(* IEC 61131-3 sources: Lasal-MCP/examples/SampleSource/LASALScreenAdvancedSolution/LASALScreenAdvancedSolution/LASALScreenAdvacnedSolution/Stations/Terminal/HMI/Class/DragDropArea, 1 file *)

(* ---- DragDropArea.st ---- *)
(*!
<Class
	Name               = "DragDropArea"
	Revision           = "0.0"
	RealtimeTask       = "false"
	CyclicTask         = "false"
	BackgroundTask     = "false"
	Sigmatek           = "false"
	OSInterface        = "false"
	HighPriority       = "false"
	Automatic          = "false"
	UpdateMode         = "Prescan"
	SharedCommandTable = "true"
	Objectsize         = "(420,240)">
	<Channels>
		<Server Name="UpdateIcon" Visualized="false" Initialize="false" WriteProtected="false" Retentive="false"/>
		<Client Name="_Grafix" Required="false" Internal="false"/>
	</Channels>
	<Network Name="DragDropArea">
		<!-- List of Components in this network -->
		<Components>
			<Object
				Name       = "_base"
				Class      = "_MyIO"
				Position   = "(218,120)"
				Visualized = "true"
				Remotely   = "true">
				<Channels>
					<Server Name="Refresh"/>
					<Server Name="Server0"/>
					<Client Name="Graphic"/>
					<Client Name="Lse"/>
				</Channels>
			</Object>
		</Components>
		<Comments>
		</Comments>
		<!-- List of Connections in this network -->
		<Connections>
			<Connection Source="this.Server0" Destination="_base.Server0" Vertices="(706,210),(534,210),"/>
			<Connection Source="this.Refresh" Destination="_base.Refresh" Vertices="(706,270),(534,270),"/>
			<Connection Source="_base.Lse" Destination="this.Lse" Vertices="(218,210),(38,210),"/>
		</Connections>
		<!-- Headerfiles -->
		<Options>
		</Options>
	</Network>
</Class>
*)
#pragma using _MyIO

DragDropArea : CLASS
: _MyIO
  //Servers:
	UpdateIcon 	: SvrCh_DINT;
  //Clients:
	_Grafix 	: CltChCmd__Grafix;
  //Variables:
		DrawClearScreen 	: BOOL;
		Started 	: BOOL;
		OnlyOnce 	: BOOL;
		SelectedLineNo 	: DINT;
		TouchCoord 	: _DOT;
		myPio 	: _IO;
		pBMP 	: ^_BMP;
  //Functions:
				//! <Function Comment="this method is called everytime when the input is active and a event occured" Name="GetEvent"/>
	FUNCTION __CDECL VIRTUAL GLOBAL GetEvent
		VAR_INPUT
			ped 	: ^_EDITOR;			//! <Variable Comment="pointer to _EDITOR information" Name="GetEvent.ped"/>
			pe 	: ^_EVENT;			//! <Variable Comment="pointer to _EVENT information" Name="GetEvent.pe"/>
		END_VAR
		VAR_OUTPUT
			retcode (EAX) 	: _DOIT;			//! <Variable Comment="for the returnstatement there are 3 different possibilities&#13;&#10;  _IDLE ..... the system should goon like it is (system goes on)&#13;&#10;  _IDIDIT ... i did it (system is ready)&#13;&#10;  _IFAILED .. i tried to do my best, but i failed (system is ready)&#13;&#10;" Name="GetEvent.retcode"/>
		END_VAR;
				//! <Function Comment="this method is called everytime when system wants to redraw the io" Name="Draw"/>
	FUNCTION __CDECL VIRTUAL GLOBAL Draw
		VAR_INPUT
			pio 	: ^_IO;			//! <Variable Comment="pointer to _IO information" Name="Draw.pio"/>
			pr 	: ^_RESULT;			//! <Variable Comment="pointer to _RESULT information" Name="Draw.pr"/>
			pv 	: ^_VARIABLE;			//! <Variable Comment="pointer to io _VARIABLE information" Name="Draw.pv"/>
			input 	: BOOL;			//! <Variable Comment="TRUE it&apos;s an input&#13;&#10;FALSE it&apos;s an output" Name="Draw.input"/>
		END_VAR
		VAR_OUTPUT
			retcode (EAX) 	: _DOIT;			//! <Variable Comment="for the returnstatement there are 3 different possibilities&#13;&#10;  _IDLE ..... the system should goon like it is (system goes on)&#13;&#10;  _IDIDIT ... i did it (system is ready)&#13;&#10;  _IFAILED .. i tried to do my best, but i failed (system is re" Name="Draw.retcode"/>
		END_VAR;

	FUNCTION GLOBAL SetIcon
		VAR_INPUT
			SelectedLine 	: DINT;
		END_VAR;

	FUNCTION GLOBAL DrawIcon
		VAR_INPUT
			CoordX 	: INT;
			CoordY 	: INT;
		END_VAR;

	FUNCTION GLOBAL DeleteIcon;

	FUNCTION GLOBAL GetDimension
		VAR_OUTPUT
			pIO 	: ^_IO;
		END_VAR;

	FUNCTION GLOBAL SetLineNo
		VAR_INPUT
			SelectedLine 	: DINT;
		END_VAR;

	FUNCTION GLOBAL ClearScreen;
  //Tables:
	FUNCTION @STD
		VAR_OUTPUT
			ret_code	: CONFSTATES;
		END_VAR;
	FUNCTION GLOBAL TAB @CT_;
END_CLASS;

#pragma usingLtd _Grafix

FUNCTION __CDECL VIRTUAL GLOBAL DragDropArea::Draw
	VAR_INPUT
		pio 	: ^_IO;
		pr 	: ^_RESULT;
		pv 	: ^_VARIABLE;
		input 	: BOOL;
	END_VAR
	VAR_OUTPUT
		retcode (EAX) 	: _DOIT;
	END_VAR
  VAR
  	act         : _NEWSCREEN;
    imageNumber : UDINT;
    myImageRoom : _ROOM;
  END_VAR

  retcode := _IDIDIT;

  _memcpy(ptr1:= #myPio, ptr2:= pio, cntr:= sizeof(myPio));

  // gets the icon once, when it is selected
  if ((Started = TRUE) & (OnlyOnce = FALSE)) then

    OnlyOnce := TRUE;

    _Grafix.GetImage(image:= #pio^.image,
                     x0:= pio^.space.xy1.x,
                     y0:= pio^.space.xy1.y,
                     x1:= pio^.space.xy2.x,
                     y1:= pio^.space.xy2.y);
  end_if;

  // returns the icon, if it is not in the IconDestList-Area
  if (DrawClearScreen = TRUE) then

    DrawClearScreen := FALSE;

    push_screen(#act);

    _Grafix.PutImage(image:= #pio^.image,
                     x0:= DEFKOORD,
                     y0:= DEFKOORD);
    pop_screen(#act);
    copy_screen(#act, #pio^.space);

  end_if;

  if (UpdateIcon = 1) then

    push_screen(#act);

    // draw background
    _Grafix.PutImage(image:= #pio^.image,
                     x0:= DEFKOORD,
                     y0:= DEFKOORD);

    imageNumber := get_no_by_label(p0:= "DragDrop",
                                   x1:= IMAGESCHEME, x2:=0);

    if (imageNumber <> DEFSCOPE) then

       pBMP$^void :=  NewDoScheme(x0:= IMAGESCHEME,
                                  x1:= SelectedLineNo,
                                  x2:= imageNumber);

      if (pBMP <> NIL) then

        myImageRoom.xy1.x := TouchCoord.x - (75/2);
        myImageRoom.xy1.y := TouchCoord.y - (75/2);
        myImageRoom.xy2.x := TouchCoord.x + (75/2);
        myImageRoom.xy2.y := TouchCoord.y + (75/2);

        out_zoom_BMP(p0:= #myImageRoom,
                     p1:= pBMP,
                     x2:= T_COPY or T_SOLID);
      end_if;
    end_if;

    pop_screen(#act);
    copy_screen(#act, #pio^.space);

  end_if;
END_FUNCTION

FUNCTION GLOBAL DragDropArea::SetIcon
	VAR_INPUT
		SelectedLine 	: DINT;
	END_VAR

  SelectedLineNo := SelectedLine;

  Started := TRUE;

END_FUNCTION

FUNCTION GLOBAL DragDropArea::DrawIcon
	VAR_INPUT
		CoordX 	: INT;
		CoordY 	: INT;
	END_VAR

  TouchCoord.x  :=  CoordX;
  TouchCoord.y  :=  CoordY;

  UpdateIcon := 1;
  Refresh := 1;

END_FUNCTION

FUNCTION GLOBAL DragDropArea::DeleteIcon

  UpdateIcon := 0;
  Started := FALSE;
  OnlyOnce := false;

END_FUNCTION

FUNCTION GLOBAL DragDropArea::GetDimension
	VAR_OUTPUT
		pIO 	: ^_IO;
	END_VAR

  pio := #myPio;

END_FUNCTION

FUNCTION GLOBAL DragDropArea::SetLineNo
	VAR_INPUT
		SelectedLine 	: DINT;
	END_VAR

  SelectedLineNo := SelectedLine;

END_FUNCTION

FUNCTION __CDECL VIRTUAL GLOBAL DragDropArea::GetEvent
	VAR_INPUT
		ped 	: ^_EDITOR;
		pe 	: ^_EVENT;
	END_VAR
	VAR_OUTPUT
		retcode (EAX) 	: _DOIT;
	END_VAR

   retcode := _MyIO::GetEvent(ped:= ped, pe:= pe);

END_FUNCTION

FUNCTION GLOBAL DragDropArea::ClearScreen

  DrawClearScreen := TRUE;
  Refresh := 1;

END_FUNCTION
